FUNCTION_BLOCK StationManager EXTENDS CyclicBase IMPLEMENTS I_StationManager
VAR
	
END_VAR

METHOD Cycle : Base_Library.HRESULT
END_METHOD

METHOD RequestNextStation : I_Station
VAR_INPUT
	CurrentStation : I_Station;
END_VAR
END_METHOD

END_FUNCTION_BLOCK

(* stored: Version 1.1.0.1
   POU StationManager: Id {418f6d70-c56b-4637-a051-e7236429bb6c}, SpecialFunc None
   Method Cycle: Id {21a5c4b4-f2de-4c1d-964f-e4b998889ed1}
   Method RequestNextStation: Id {0f9d2668-e50b-4e8a-9785-225d9d2f5583} *)
